FUNCTION_BLOCK Subestacao_HMI (* Service Interface Function Block Type *)
  (* Standard: 61499-2 *)
  (* Version 1.1, 15/10/2026, Hidryco, Hidryco, Hidryco 04/11/2026: comandos ABRIR_/FECHAR_1Qx gravaveis como no legado (um evento por comando); pulso na bobina = PULSO_ABRIR_/PULSO_FECHAR_1Qx. Nomes do legado (Unifilar): LOCAL_/REMOTO_/PRONTO_/CARREGADO_/SEM_FALHA_1Qx (eram MPL_/MPR_/MPP_/MPC_/MPSF_), ABRIR_/FECHAR_1Qx (eram CMD_ABRIR/CMD_FECHAR1Qx) e novas ABERTO_/FECHADO_1Qx. IHM da Subestacao (unifilar do QGBT e cargas no gerador) *)
  PACKAGE Hidryco.HidrycoLib;
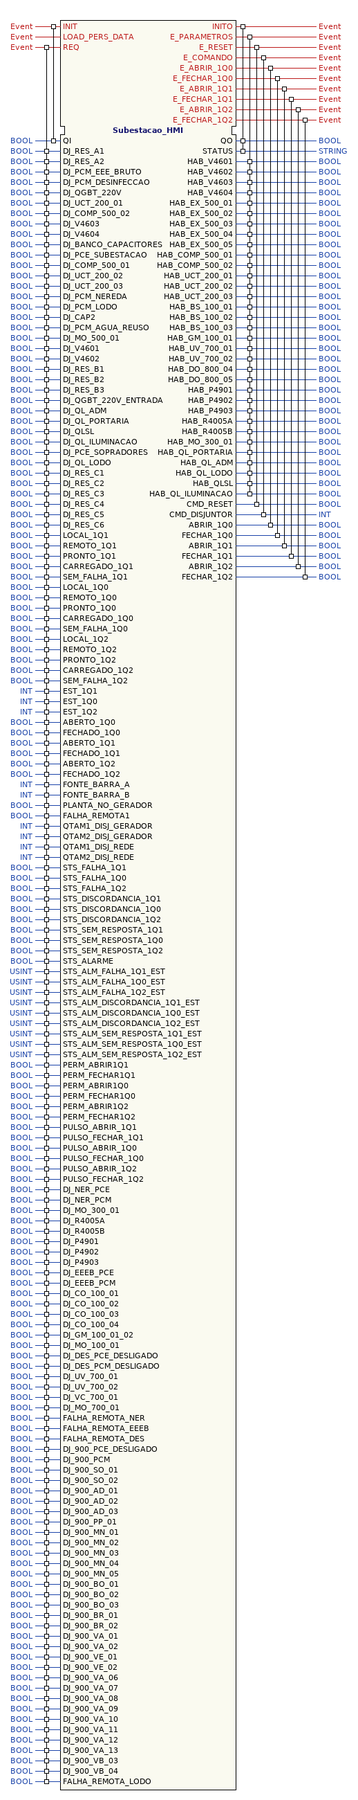
  EVENT_INPUT
    INIT WITH QI;
    LOAD_PERS_DATA; (* Reenvia os parametros persistentes *)
    REQ WITH DJ_RES_A1, DJ_RES_A2, DJ_PCM_EEE_BRUTO, DJ_PCM_DESINFECCAO, DJ_QGBT_220V, DJ_UCT_200_01, DJ_COMP_500_02, DJ_V4603, DJ_V4604, DJ_BANCO_CAPACITORES, DJ_PCE_SUBESTACAO, DJ_COMP_500_01, DJ_UCT_200_02, DJ_UCT_200_03, DJ_PCM_NEREDA, DJ_PCM_LODO, DJ_CAP2, DJ_PCM_AGUA_REUSO, DJ_MO_500_01, DJ_V4601, DJ_V4602, DJ_RES_B1, DJ_RES_B2, DJ_RES_B3, DJ_QGBT_220V_ENTRADA, DJ_QL_ADM, DJ_QL_PORTARIA, DJ_QLSL, DJ_QL_ILUMINACAO, DJ_PCE_SOPRADORES, DJ_QL_LODO, DJ_RES_C1, DJ_RES_C2, DJ_RES_C3, DJ_RES_C4, DJ_RES_C5, DJ_RES_C6, LOCAL_1Q1, REMOTO_1Q1, PRONTO_1Q1, CARREGADO_1Q1, SEM_FALHA_1Q1, LOCAL_1Q0, REMOTO_1Q0, PRONTO_1Q0, CARREGADO_1Q0, SEM_FALHA_1Q0, LOCAL_1Q2, REMOTO_1Q2, PRONTO_1Q2, CARREGADO_1Q2, SEM_FALHA_1Q2, EST_1Q1, EST_1Q0, EST_1Q2, FONTE_BARRA_A, FONTE_BARRA_B, PLANTA_NO_GERADOR, FALHA_REMOTA1, QTAM1_DISJ_GERADOR, QTAM2_DISJ_GERADOR, QTAM1_DISJ_REDE, QTAM2_DISJ_REDE, STS_FALHA_1Q1, STS_FALHA_1Q0, STS_FALHA_1Q2, STS_DISCORDANCIA_1Q1, STS_DISCORDANCIA_1Q0, STS_DISCORDANCIA_1Q2, STS_SEM_RESPOSTA_1Q1, STS_SEM_RESPOSTA_1Q0, STS_SEM_RESPOSTA_1Q2, STS_ALARME, STS_ALM_FALHA_1Q1_EST, STS_ALM_FALHA_1Q0_EST, STS_ALM_FALHA_1Q2_EST, STS_ALM_DISCORDANCIA_1Q1_EST, STS_ALM_DISCORDANCIA_1Q0_EST, STS_ALM_DISCORDANCIA_1Q2_EST, STS_ALM_SEM_RESPOSTA_1Q1_EST, STS_ALM_SEM_RESPOSTA_1Q0_EST, STS_ALM_SEM_RESPOSTA_1Q2_EST, PERM_ABRIR1Q1, PERM_FECHAR1Q1, PERM_ABRIR1Q0, PERM_FECHAR1Q0, PERM_ABRIR1Q2, PERM_FECHAR1Q2, PULSO_ABRIR_1Q1, PULSO_FECHAR_1Q1, PULSO_ABRIR_1Q0, PULSO_FECHAR_1Q0, PULSO_ABRIR_1Q2, PULSO_FECHAR_1Q2, DJ_NER_PCE, DJ_NER_PCM, DJ_MO_300_01, DJ_R4005A, DJ_R4005B, DJ_P4901, DJ_P4902, DJ_P4903, DJ_EEEB_PCE, DJ_EEEB_PCM, DJ_CO_100_01, DJ_CO_100_02, DJ_CO_100_03, DJ_CO_100_04, DJ_GM_100_01_02, DJ_MO_100_01, DJ_DES_PCE_DESLIGADO, DJ_DES_PCM_DESLIGADO, DJ_UV_700_01, DJ_UV_700_02, DJ_VC_700_01, DJ_MO_700_01, FALHA_REMOTA_NER, FALHA_REMOTA_EEEB, FALHA_REMOTA_DES, ABERTO_1Q0, FECHADO_1Q0, ABERTO_1Q1, FECHADO_1Q1, ABERTO_1Q2, FECHADO_1Q2, DJ_900_PCE_DESLIGADO, DJ_900_PCM, DJ_900_SO_01, DJ_900_SO_02, DJ_900_AD_01, DJ_900_AD_02, DJ_900_AD_03, DJ_900_PP_01, DJ_900_MN_01, DJ_900_MN_02, DJ_900_MN_03, DJ_900_MN_04, DJ_900_MN_05, DJ_900_BO_01, DJ_900_BO_02, DJ_900_BO_03, DJ_900_BR_01, DJ_900_BR_02, DJ_900_VA_01, DJ_900_VA_02, DJ_900_VE_01, DJ_900_VE_02, DJ_900_VA_06, DJ_900_VA_07, DJ_900_VA_08, DJ_900_VA_09, DJ_900_VA_10, DJ_900_VA_11, DJ_900_VA_12, DJ_900_VA_13, DJ_900_VB_03, DJ_900_VB_04, FALHA_REMOTA_LODO; (* Atualizacao de status *)
  END_EVENT
  EVENT_OUTPUT
    INITO WITH QO, STATUS;
    E_PARAMETROS WITH HAB_V4601, HAB_V4602, HAB_V4603, HAB_V4604, HAB_EX_500_01, HAB_EX_500_02, HAB_EX_500_03, HAB_EX_500_04, HAB_EX_500_05, HAB_COMP_500_01, HAB_COMP_500_02, HAB_UCT_200_01, HAB_UCT_200_02, HAB_UCT_200_03, HAB_BS_100_01, HAB_BS_100_02, HAB_BS_100_03, HAB_GM_100_01, HAB_UV_700_01, HAB_UV_700_02, HAB_DO_800_04, HAB_DO_800_05, HAB_P4901, HAB_P4902, HAB_P4903, HAB_R4005A, HAB_R4005B, HAB_MO_300_01, HAB_QL_PORTARIA, HAB_QL_ADM, HAB_QL_LODO, HAB_QLSL, HAB_QL_ILUMINACAO;
    E_RESET WITH CMD_RESET;
    E_COMANDO WITH CMD_DISJUNTOR;
    E_ABRIR_1Q0 WITH ABRIR_1Q0; (* Comando ABRIR_1Q0 (como no legado): TRUE = executa *)
    E_FECHAR_1Q0 WITH FECHAR_1Q0; (* Comando FECHAR_1Q0 (como no legado): TRUE = executa *)
    E_ABRIR_1Q1 WITH ABRIR_1Q1; (* Comando ABRIR_1Q1 (como no legado): TRUE = executa *)
    E_FECHAR_1Q1 WITH FECHAR_1Q1; (* Comando FECHAR_1Q1 (como no legado): TRUE = executa *)
    E_ABRIR_1Q2 WITH ABRIR_1Q2; (* Comando ABRIR_1Q2 (como no legado): TRUE = executa *)
    E_FECHAR_1Q2 WITH FECHAR_1Q2; (* Comando FECHAR_1Q2 (como no legado): TRUE = executa *)
  END_EVENT
  VAR_INPUT
    QI : BOOL;
    DJ_RES_A1 : BOOL; (* Disjuntor RES_A1 ligado *)
    DJ_RES_A2 : BOOL; (* Disjuntor RES_A2 ligado *)
    DJ_PCM_EEE_BRUTO : BOOL; (* Disjuntor PCM_EEE_BRUTO ligado *)
    DJ_PCM_DESINFECCAO : BOOL; (* Disjuntor PCM_DESINFECCAO ligado *)
    DJ_QGBT_220V : BOOL; (* Disjuntor QGBT_220V ligado *)
    DJ_UCT_200_01 : BOOL; (* Disjuntor UCT_200_01 ligado *)
    DJ_COMP_500_02 : BOOL; (* Disjuntor COMP_500_02 ligado *)
    DJ_V4603 : BOOL; (* Disjuntor V4603 ligado *)
    DJ_V4604 : BOOL; (* Disjuntor V4604 ligado *)
    DJ_BANCO_CAPACITORES : BOOL; (* Disjuntor BANCO_CAPACITORES ligado *)
    DJ_PCE_SUBESTACAO : BOOL; (* Disjuntor PCE_SUBESTACAO ligado *)
    DJ_COMP_500_01 : BOOL; (* Disjuntor COMP_500_01 ligado *)
    DJ_UCT_200_02 : BOOL; (* Disjuntor UCT_200_02 ligado *)
    DJ_UCT_200_03 : BOOL; (* Disjuntor UCT_200_03 ligado *)
    DJ_PCM_NEREDA : BOOL; (* Disjuntor PCM_NEREDA ligado *)
    DJ_PCM_LODO : BOOL; (* Disjuntor PCM_LODO ligado *)
    DJ_CAP2 : BOOL; (* Disjuntor CAP2 ligado *)
    DJ_PCM_AGUA_REUSO : BOOL; (* Disjuntor PCM_AGUA_REUSO ligado *)
    DJ_MO_500_01 : BOOL; (* Disjuntor MO_500_01 ligado *)
    DJ_V4601 : BOOL; (* Disjuntor V4601 ligado *)
    DJ_V4602 : BOOL; (* Disjuntor V4602 ligado *)
    DJ_RES_B1 : BOOL; (* Disjuntor RES_B1 ligado *)
    DJ_RES_B2 : BOOL; (* Disjuntor RES_B2 ligado *)
    DJ_RES_B3 : BOOL; (* Disjuntor RES_B3 ligado *)
    DJ_QGBT_220V_ENTRADA : BOOL; (* Disjuntor QGBT_220V_ENTRADA ligado *)
    DJ_QL_ADM : BOOL; (* Disjuntor QL_ADM ligado *)
    DJ_QL_PORTARIA : BOOL; (* Disjuntor QL_PORTARIA ligado *)
    DJ_QLSL : BOOL; (* Disjuntor QLSL ligado *)
    DJ_QL_ILUMINACAO : BOOL; (* Disjuntor QL_ILUMINACAO ligado *)
    DJ_PCE_SOPRADORES : BOOL; (* Disjuntor PCE_SOPRADORES ligado *)
    DJ_QL_LODO : BOOL; (* Disjuntor QL_LODO ligado *)
    DJ_RES_C1 : BOOL; (* Disjuntor RES_C1 ligado *)
    DJ_RES_C2 : BOOL; (* Disjuntor RES_C2 ligado *)
    DJ_RES_C3 : BOOL; (* Disjuntor RES_C3 ligado *)
    DJ_RES_C4 : BOOL; (* Disjuntor RES_C4 ligado *)
    DJ_RES_C5 : BOOL; (* Disjuntor RES_C5 ligado *)
    DJ_RES_C6 : BOOL; (* Disjuntor RES_C6 ligado *)
    LOCAL_1Q1 : BOOL; (* Local 1Q1 *)
    REMOTO_1Q1 : BOOL; (* Remoto 1Q1 *)
    PRONTO_1Q1 : BOOL; (* Pronto para fechar 1Q1 *)
    CARREGADO_1Q1 : BOOL; (* Mola carregada 1Q1 *)
    SEM_FALHA_1Q1 : BOOL; (* Sem falha 1Q1 *)
    LOCAL_1Q0 : BOOL; (* Local 1Q0 *)
    REMOTO_1Q0 : BOOL; (* Remoto 1Q0 *)
    PRONTO_1Q0 : BOOL; (* Pronto para fechar 1Q0 *)
    CARREGADO_1Q0 : BOOL; (* Mola carregada 1Q0 *)
    SEM_FALHA_1Q0 : BOOL; (* Sem falha 1Q0 *)
    LOCAL_1Q2 : BOOL; (* Local 1Q2 *)
    REMOTO_1Q2 : BOOL; (* Remoto 1Q2 *)
    PRONTO_1Q2 : BOOL; (* Pronto para fechar 1Q2 *)
    CARREGADO_1Q2 : BOOL; (* Mola carregada 1Q2 *)
    SEM_FALHA_1Q2 : BOOL; (* Sem falha 1Q2 *)
    EST_1Q1 : INT; (* Disjuntor 1Q1: 0 indefinido (sem comunicacao), 1 aberto, 2 fechado, 3 discordante *)
    EST_1Q0 : INT; (* Disjuntor 1Q0: 0 indefinido (sem comunicacao), 1 aberto, 2 fechado, 3 discordante *)
    EST_1Q2 : INT; (* Disjuntor 1Q2: 0 indefinido (sem comunicacao), 1 aberto, 2 fechado, 3 discordante *)
    ABERTO_1Q0 : BOOL; (* Disjuntor 1Q0 aberto (contato do campo) *)
    FECHADO_1Q0 : BOOL; (* Disjuntor 1Q0 fechado (contato do campo) *)
    ABERTO_1Q1 : BOOL; (* Disjuntor 1Q1 aberto (contato do campo) *)
    FECHADO_1Q1 : BOOL; (* Disjuntor 1Q1 fechado (contato do campo) *)
    ABERTO_1Q2 : BOOL; (* Disjuntor 1Q2 aberto (contato do campo) *)
    FECHADO_1Q2 : BOOL; (* Disjuntor 1Q2 fechado (contato do campo) *)
    FONTE_BARRA_A : INT; (* Fonte da barra A (1Q1): 0 sem alimentacao, 1 rede, 2 gerador, 3 indefinida *)
    FONTE_BARRA_B : INT; (* Fonte da barra B (1Q2): 0 sem alimentacao, 1 rede, 2 gerador, 3 indefinida *)
    PLANTA_NO_GERADOR : BOOL; (* Alguma QTAM com o disjuntor do gerador fechado (planta nos geradores) *)
    FALHA_REMOTA1 : BOOL; (* Falha de comunicacao com a remota 1 *)
    QTAM1_DISJ_GERADOR : INT; (* QTAM1: disjuntor do gerador G2 (0 indef., 1 aberto, 2 fechado) *)
    QTAM2_DISJ_GERADOR : INT; (* QTAM2: disjuntor do gerador G1 (0 indef., 1 aberto, 2 fechado) *)
    QTAM1_DISJ_REDE : INT; (* QTAM1: disjuntor de rede (0 indef., 1 aberto, 2 fechado) *)
    QTAM2_DISJ_REDE : INT; (* QTAM2: disjuntor de rede (0 indef., 1 aberto, 2 fechado) *)
    STS_FALHA_1Q1 : BOOL; (* Disjuntor 1Q1 em falha (desarmado) *)
    STS_FALHA_1Q0 : BOOL; (* Disjuntor 1Q0 em falha (desarmado) *)
    STS_FALHA_1Q2 : BOOL; (* Disjuntor 1Q2 em falha (desarmado) *)
    STS_DISCORDANCIA_1Q1 : BOOL; (* Disjuntor 1Q1: posição indefinida (aberto e fechado discordantes) *)
    STS_DISCORDANCIA_1Q0 : BOOL; (* Disjuntor 1Q0: posição indefinida (aberto e fechado discordantes) *)
    STS_DISCORDANCIA_1Q2 : BOOL; (* Disjuntor 1Q2: posição indefinida (aberto e fechado discordantes) *)
    STS_SEM_RESPOSTA_1Q1 : BOOL; (* Disjuntor 1Q1 não respondeu ao comando de abrir/fechar *)
    STS_SEM_RESPOSTA_1Q0 : BOOL; (* Disjuntor 1Q0 não respondeu ao comando de abrir/fechar *)
    STS_SEM_RESPOSTA_1Q2 : BOOL; (* Disjuntor 1Q2 não respondeu ao comando de abrir/fechar *)
    STS_ALARME : BOOL; (* Algum alarme do QGBT *)
    STS_ALM_FALHA_1Q1_EST : USINT; (* Estado do ALARM_BIT Disjuntor 1Q1 em falha (desarmado) (0 normal, 1 ativo reconhecido, 2 ativo nao reconhecido, 3 saiu nao reconhecido, 4 ativo e saiu nao reconhecido) *)
    STS_ALM_FALHA_1Q0_EST : USINT; (* Estado do ALARM_BIT Disjuntor 1Q0 em falha (desarmado) (0 normal, 1 ativo reconhecido, 2 ativo nao reconhecido, 3 saiu nao reconhecido, 4 ativo e saiu nao reconhecido) *)
    STS_ALM_FALHA_1Q2_EST : USINT; (* Estado do ALARM_BIT Disjuntor 1Q2 em falha (desarmado) (0 normal, 1 ativo reconhecido, 2 ativo nao reconhecido, 3 saiu nao reconhecido, 4 ativo e saiu nao reconhecido) *)
    STS_ALM_DISCORDANCIA_1Q1_EST : USINT; (* Estado do ALARM_BIT Disjuntor 1Q1: posição indefinida (aberto e fechado discordantes) (0 normal, 1 ativo reconhecido, 2 ativo nao reconhecido, 3 saiu nao reconhecido, 4 ativo e saiu nao reconhecido) *)
    STS_ALM_DISCORDANCIA_1Q0_EST : USINT; (* Estado do ALARM_BIT Disjuntor 1Q0: posição indefinida (aberto e fechado discordantes) (0 normal, 1 ativo reconhecido, 2 ativo nao reconhecido, 3 saiu nao reconhecido, 4 ativo e saiu nao reconhecido) *)
    STS_ALM_DISCORDANCIA_1Q2_EST : USINT; (* Estado do ALARM_BIT Disjuntor 1Q2: posição indefinida (aberto e fechado discordantes) (0 normal, 1 ativo reconhecido, 2 ativo nao reconhecido, 3 saiu nao reconhecido, 4 ativo e saiu nao reconhecido) *)
    STS_ALM_SEM_RESPOSTA_1Q1_EST : USINT; (* Estado do ALARM_BIT Disjuntor 1Q1 não respondeu ao comando de abrir/fechar (0 normal, 1 ativo reconhecido, 2 ativo nao reconhecido, 3 saiu nao reconhecido, 4 ativo e saiu nao reconhecido) *)
    STS_ALM_SEM_RESPOSTA_1Q0_EST : USINT; (* Estado do ALARM_BIT Disjuntor 1Q0 não respondeu ao comando de abrir/fechar (0 normal, 1 ativo reconhecido, 2 ativo nao reconhecido, 3 saiu nao reconhecido, 4 ativo e saiu nao reconhecido) *)
    STS_ALM_SEM_RESPOSTA_1Q2_EST : USINT; (* Estado do ALARM_BIT Disjuntor 1Q2 não respondeu ao comando de abrir/fechar (0 normal, 1 ativo reconhecido, 2 ativo nao reconhecido, 3 saiu nao reconhecido, 4 ativo e saiu nao reconhecido) *)
    PERM_ABRIR1Q1 : BOOL; (* IHM: abrir o 1Q1 permitido *)
    PERM_FECHAR1Q1 : BOOL; (* IHM: fechar o 1Q1 permitido *)
    PERM_ABRIR1Q0 : BOOL; (* IHM: abrir o 1Q0 permitido *)
    PERM_FECHAR1Q0 : BOOL; (* IHM: fechar o 1Q0 permitido *)
    PERM_ABRIR1Q2 : BOOL; (* IHM: abrir o 1Q2 permitido *)
    PERM_FECHAR1Q2 : BOOL; (* IHM: fechar o 1Q2 permitido *)
    PULSO_ABRIR_1Q1 : BOOL; (* Pulso de abrir o 1Q1 (bobina MX) *)
    PULSO_FECHAR_1Q1 : BOOL; (* Pulso de fechar o 1Q1 (bobina XF) *)
    PULSO_ABRIR_1Q0 : BOOL; (* Pulso de abrir o 1Q0 (bobina MX) *)
    PULSO_FECHAR_1Q0 : BOOL; (* Pulso de fechar o 1Q0 (bobina XF) *)
    PULSO_ABRIR_1Q2 : BOOL; (* Pulso de abrir o 1Q2 (bobina MX) *)
    PULSO_FECHAR_1Q2 : BOOL; (* Pulso de fechar o 1Q2 (bobina XF) *)
    DJ_NER_PCE : BOOL; (* Painel Nereda: disjuntor PCE ligado (remota Nereda A3 %I0.0) *)
    DJ_NER_PCM : BOOL; (* Painel Nereda: disjuntor PCM Nereda ligado (A3 %I0.2) *)
    DJ_MO_300_01 : BOOL; (* Painel Nereda: disjuntor 300-MO-01 ligado (A3 %I0.6) *)
    DJ_R4005A : BOOL; (* Painel Nereda: disjuntor R4005A ligado (A3 %I0.22) *)
    DJ_R4005B : BOOL; (* Painel Nereda: disjuntor R4005B ligado (A3 %I0.23) *)
    DJ_P4901 : BOOL; (* Painel Nereda: disjuntor P4901 ligado (A4 %I0.34) *)
    DJ_P4902 : BOOL; (* Painel Nereda: disjuntor P4902 ligado (A4 %I0.35) *)
    DJ_P4903 : BOOL; (* Painel Nereda: disjuntor P4903 ligado (A4 %I0.36) *)
    DJ_EEEB_PCE : BOOL; (* Painel EEE Bruto: disjuntor PCE ligado (remota EEE A2 %I0.0) *)
    DJ_EEEB_PCM : BOOL; (* Painel EEE Bruto: disjuntor PCM EEE Bruto ligado (A2 %I0.2) *)
    DJ_CO_100_01 : BOOL; (* Painel EEE Bruto: disjuntor 100-CO-01 ligado (A2 %I0.6) *)
    DJ_CO_100_02 : BOOL; (* Painel EEE Bruto: disjuntor 100-CO-02 ligado (A2 %I0.7) *)
    DJ_CO_100_03 : BOOL; (* Painel EEE Bruto: disjuntor 100-CO-03 ligado (A2 %I0.8) *)
    DJ_CO_100_04 : BOOL; (* Painel EEE Bruto: disjuntor 100-CO-04 ligado (A2 %I0.9) *)
    DJ_GM_100_01_02 : BOOL; (* Painel EEE Bruto: disjuntor 100-GM-01/02 ligado (A2 %I0.10) *)
    DJ_MO_100_01 : BOOL; (* Painel EEE Bruto: disjuntor 100-MO-01 ligado (A2 %I0.11) *)
    DJ_DES_PCE_DESLIGADO : BOOL; (* Painel Desinfeccao: disjuntor PCE DESLIGADO (remota Desinfeccao A2 %I0.0, logica invertida) *)
    DJ_DES_PCM_DESLIGADO : BOOL; (* Painel Desinfeccao: disjuntor PCM DESLIGADO (A2 %I0.1, logica invertida) *)
    DJ_UV_700_01 : BOOL; (* Painel Desinfeccao: disjuntor 700-UV-01 ligado (A2 %I0.2) *)
    DJ_UV_700_02 : BOOL; (* Painel Desinfeccao: disjuntor 700-UV-02 ligado (A2 %I0.3) *)
    DJ_VC_700_01 : BOOL; (* Painel Desinfeccao: disjuntor 700-VC-01 ligado (A2 %I0.4) *)
    DJ_MO_700_01 : BOOL; (* Painel Desinfeccao: disjuntor 700-MO-01 ligado (A2 %I0.5) *)
    FALHA_REMOTA_NER : BOOL; (* Falha de comunicacao do M262_Substacao com a remota 1 Nereda (10.26.208.160) *)
    FALHA_REMOTA_EEEB : BOOL; (* Falha de comunicacao do M262_Substacao com a remota EEE Bruto (10.26.208.197) *)
    FALHA_REMOTA_DES : BOOL; (* Falha de comunicacao do M262_Substacao com a remota Desinfeccao (10.26.208.137) *)
    DJ_900_PCE_DESLIGADO : BOOL; (* Painel Lodo (PCE LODO 900): disjuntor PCE DESLIGADO (remota Lodo .135 A3 %I0.0, logica invertida) *)
    DJ_900_PCM : BOOL; (* Painel Lodo (PCE LODO 900): disjuntor PCM ligado (remota Lodo .135 A3 %I0.2) *)
    DJ_900_SO_01 : BOOL; (* Painel Lodo (PCE LODO 900): disjuntor SO-01 ligado (remota Lodo .135 A3 %I0.3) *)
    DJ_900_SO_02 : BOOL; (* Painel Lodo (PCE LODO 900): disjuntor SO-02 ligado (remota Lodo .135 A3 %I0.8) *)
    DJ_900_AD_01 : BOOL; (* Painel Lodo (PCE LODO 900): disjuntor AD-01 ligado (remota Lodo .135 A3 %I0.13) *)
    DJ_900_AD_02 : BOOL; (* Painel Lodo (PCE LODO 900): disjuntor AD-02 ligado (remota Lodo .135 A3 %I0.14) *)
    DJ_900_AD_03 : BOOL; (* Painel Lodo (PCE LODO 900): disjuntor AD-03 ligado (remota Lodo .135 A3 %I0.15) *)
    DJ_900_PP_01 : BOOL; (* Painel Lodo (PCE LODO 900): disjuntor PP-01 ligado (remota Lodo .135 A3 %I0.16) *)
    DJ_900_MN_01 : BOOL; (* Painel Lodo (PCE LODO 900): disjuntor MN-01 ligado (remota Lodo .135 A3 %I0.17) *)
    DJ_900_MN_02 : BOOL; (* Painel Lodo (PCE LODO 900): disjuntor MN-02 ligado (remota Lodo .135 A3 %I0.18) *)
    DJ_900_MN_03 : BOOL; (* Painel Lodo (PCE LODO 900): disjuntor MN-03 ligado (remota Lodo .135 A3 %I0.19) *)
    DJ_900_MN_04 : BOOL; (* Painel Lodo (PCE LODO 900): disjuntor MN-04 ligado (remota Lodo .135 A3 %I0.20) *)
    DJ_900_MN_05 : BOOL; (* Painel Lodo (PCE LODO 900): disjuntor MN-05 ligado (remota Lodo .135 A3 %I0.21) *)
    DJ_900_BO_01 : BOOL; (* Painel Lodo (PCE LODO 900): disjuntor BO-01 ligado (remota Lodo .135 A3 %I0.22) *)
    DJ_900_BO_02 : BOOL; (* Painel Lodo (PCE LODO 900): disjuntor BO-02 ligado (remota Lodo .135 A3 %I0.28) *)
    DJ_900_BO_03 : BOOL; (* Painel Lodo (PCE LODO 900): disjuntor BO-03 ligado (remota Lodo .135 A4 %I0.34) *)
    DJ_900_BR_01 : BOOL; (* Painel Lodo (PCE LODO 900): disjuntor BR-01 ligado (remota Lodo .135 A4 %I0.40) *)
    DJ_900_BR_02 : BOOL; (* Painel Lodo (PCE LODO 900): disjuntor BR-02 ligado (remota Lodo .135 A4 %I0.46) *)
    DJ_900_VA_01 : BOOL; (* Painel Lodo (PCE LODO 900): disjuntor VA-01 ligado (remota Lodo .135 A4 %I0.52) *)
    DJ_900_VA_02 : BOOL; (* Painel Lodo (PCE LODO 900): disjuntor VA-02 ligado (remota Lodo .135 A4 %I0.53) *)
    DJ_900_VE_01 : BOOL; (* Painel Lodo (PCE LODO 900): disjuntor VE-01 ligado (remota Lodo .135 A4 %I0.54) *)
    DJ_900_VE_02 : BOOL; (* Painel Lodo (PCE LODO 900): disjuntor VE-02 ligado (remota Lodo .135 A4 %I0.55) *)
    DJ_900_VA_06 : BOOL; (* Painel Lodo (PCE LODO 900): disjuntor VA-06 ligado (remota Lodo .135 A4 %I0.57) *)
    DJ_900_VA_07 : BOOL; (* Painel Lodo (PCE LODO 900): disjuntor VA-07 ligado (remota Lodo .135 A4 %I0.58) *)
    DJ_900_VA_08 : BOOL; (* Painel Lodo (PCE LODO 900): disjuntor VA-08 ligado (remota Lodo .135 A4 %I0.59) *)
    DJ_900_VA_09 : BOOL; (* Painel Lodo (PCE LODO 900): disjuntor VA-09 ligado (remota Lodo .135 A4 %I0.60) *)
    DJ_900_VA_10 : BOOL; (* Painel Lodo (PCE LODO 900): disjuntor VA-10 ligado (remota Lodo .135 A4 %I0.61) *)
    DJ_900_VA_11 : BOOL; (* Painel Lodo (PCE LODO 900): disjuntor VA-11 ligado (remota Lodo .135 A4 %I0.62) *)
    DJ_900_VA_12 : BOOL; (* Painel Lodo (PCE LODO 900): disjuntor VA-12 ligado (remota Lodo .135 A4 %I0.63) *)
    DJ_900_VA_13 : BOOL; (* Painel Lodo (PCE LODO 900): disjuntor VA-13 ligado (remota Lodo .135 A5 %I0.64) *)
    DJ_900_VB_03 : BOOL; (* Painel Lodo (PCE LODO 900): disjuntor VB-03 ligado (remota Lodo .135 A5 %I0.65) *)
    DJ_900_VB_04 : BOOL; (* Painel Lodo (PCE LODO 900): disjuntor VB-04 ligado (remota Lodo .135 A5 %I0.66) *)
    FALHA_REMOTA_LODO : BOOL; (* Falha de comunicacao do M262_Substacao com a remota 1 do PCE LODO (10.26.208.135) *)
  END_VAR
  VAR_OUTPUT
    QO : BOOL; (* Event Output Qualifier *)
    STATUS : STRING; (* Service Status *)
    HAB_V4601 : BOOL; (* V4601 - Soprador 01 liberado com a planta nos geradores *)
    HAB_V4602 : BOOL; (* V4602 - Soprador 02 liberado com a planta nos geradores *)
    HAB_V4603 : BOOL; (* V4603 - Soprador 03 liberado com a planta nos geradores *)
    HAB_V4604 : BOOL; (* V4604 - Soprador 04 liberado com a planta nos geradores *)
    HAB_EX_500_01 : BOOL; (* 500-EX-01 - Exaustor 01 liberado com a planta nos geradores *)
    HAB_EX_500_02 : BOOL; (* 500-EX-02 - Exaustor 02 liberado com a planta nos geradores *)
    HAB_EX_500_03 : BOOL; (* 500-EX-03 - Exaustor 03 liberado com a planta nos geradores *)
    HAB_EX_500_04 : BOOL; (* 500-EX-04 - Exaustor 04 liberado com a planta nos geradores *)
    HAB_EX_500_05 : BOOL; (* 500-EX-05 - Exaustor 05 liberado com a planta nos geradores *)
    HAB_COMP_500_01 : BOOL; (* 500-COMP-01 - Compressor 01 liberado com a planta nos geradores *)
    HAB_COMP_500_02 : BOOL; (* 500-COMP-02 - Compressor 02 liberado com a planta nos geradores *)
    HAB_UCT_200_01 : BOOL; (* 200-UCT-01 - Unid. compacta 01 liberado com a planta nos geradores *)
    HAB_UCT_200_02 : BOOL; (* 200-UCT-02 - Unid. compacta 02 liberado com a planta nos geradores *)
    HAB_UCT_200_03 : BOOL; (* 200-UCT-03 - Unid. compacta 03 liberado com a planta nos geradores *)
    HAB_BS_100_01 : BOOL; (* 100-BS-01 - Bomba 01 liberado com a planta nos geradores *)
    HAB_BS_100_02 : BOOL; (* 100-BS-02 - Bomba 02 liberado com a planta nos geradores *)
    HAB_BS_100_03 : BOOL; (* 100-BS-03 - Bomba 03 liberado com a planta nos geradores *)
    HAB_GM_100_01 : BOOL; (* 100-GM-01 - Grade mecanizada liberado com a planta nos geradores *)
    HAB_UV_700_01 : BOOL; (* 700-UV-01 - Sistema UV 01 liberado com a planta nos geradores *)
    HAB_UV_700_02 : BOOL; (* 700-UV-02 - Sistema UV 02 liberado com a planta nos geradores *)
    HAB_DO_800_04 : BOOL; (* 800-DO-04 - Bomba dosadora 04 liberado com a planta nos geradores *)
    HAB_DO_800_05 : BOOL; (* 800-DO-05 - Bomba dosadora 05 liberado com a planta nos geradores *)
    HAB_P4901 : BOOL; (* P4901 - Bomba submersível 01 liberado com a planta nos geradores *)
    HAB_P4902 : BOOL; (* P4902 - Bomba submersível 02 liberado com a planta nos geradores *)
    HAB_P4903 : BOOL; (* P4903 - Bomba submersível 03 liberado com a planta nos geradores *)
    HAB_R4005A : BOOL; (* R4005A - Bomba horizontal A liberado com a planta nos geradores *)
    HAB_R4005B : BOOL; (* R4005B - Bomba horizontal B liberado com a planta nos geradores *)
    HAB_MO_300_01 : BOOL; (* 300-MO-01 - Misturador 01 liberado com a planta nos geradores *)
    HAB_QL_PORTARIA : BOOL; (* QL Portaria liberado com a planta nos geradores *)
    HAB_QL_ADM : BOOL; (* QL Administração liberado com a planta nos geradores *)
    HAB_QL_LODO : BOOL; (* QL Lodo liberado com a planta nos geradores *)
    HAB_QLSL : BOOL; (* QL Sala de quadros liberado com a planta nos geradores *)
    HAB_QL_ILUMINACAO : BOOL; (* QL Iluminação externa liberado com a planta nos geradores *)
    CMD_RESET : BOOL; (* Reconhece os alarmes do QGBT e dos geradores *)
    CMD_DISJUNTOR : INT; (* Comando dos Masterpact: 1/2 abrir/fechar 1Q1, 3/4 abrir/fechar 1Q0, 5/6 abrir/fechar 1Q2 *)
    ABRIR_1Q0 : BOOL; (* Comando abrir do disjuntor 1Q0 (legado): TRUE = executa, com as mesmas permissoes do faceplate *)
    FECHAR_1Q0 : BOOL; (* Comando fechar do disjuntor 1Q0 (legado): TRUE = executa, com as mesmas permissoes do faceplate *)
    ABRIR_1Q1 : BOOL; (* Comando abrir do disjuntor 1Q1 (legado): TRUE = executa, com as mesmas permissoes do faceplate *)
    FECHAR_1Q1 : BOOL; (* Comando fechar do disjuntor 1Q1 (legado): TRUE = executa, com as mesmas permissoes do faceplate *)
    ABRIR_1Q2 : BOOL; (* Comando abrir do disjuntor 1Q2 (legado): TRUE = executa, com as mesmas permissoes do faceplate *)
    FECHAR_1Q2 : BOOL; (* Comando fechar do disjuntor 1Q2 (legado): TRUE = executa, com as mesmas permissoes do faceplate *)
  END_VAR
  SERVICE /
    SEQUENCE 
    END_SEQUENCE
  END_SERVICE
END_FUNCTION_BLOCK
